ADAPTER IWorkpieceSupply (* Adapter Interface *)
  (* Standard: 61499-1 *)
  (* Version 0.0, 11/16/2026, Sandeep Patil, Flexbridge AB *)
  PACKAGE Flexbridge.FestoMPS400;
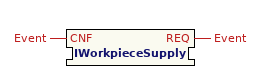
  EVENT_INPUT
    CNF; (* To the plug: the workpiece has been handed over *)
  END_EVENT
  EVENT_OUTPUT
    REQ; (* From the plug: please hand over one workpiece *)
  END_EVENT
  SERVICE SOCKET/PLUG
    SEQUENCE request_workpiece
      PLUG.REQ() -> SOCKET.REQ();
      SOCKET.CNF() -> PLUG.CNF();
    END_SEQUENCE
  END_SERVICE
END_ADAPTER
